// TIA Portal V20 export
DATA_BLOCK "DB_DATA_LASER"   // DB401
{ S7_Optimized_Access := 'TRUE' }
// stored: AutoNumber false, MemoryReserve 100
   VAR
      LASER_DATA_READ : Array[0..71] of Byte;
      LASER_DATA_WRITE : Array[0..71] of Byte;
      READ : Bool;
      WRITE : Bool;
   END_VAR
BEGIN
END_DATA_BLOCK
